// TIA Portal V17 program export: 0 tag tables, 0 data types, 1 data blocks, 1 code blocks (in call order from the OBs), 0 instance data blocks

DATA_BLOCK "流水灯定时器"   // DB1
{ S7_Optimized_Access := 'FALSE' }
   VAR
      黄灯计时 : TON_TIME;
      蓝灯计时 : TON_TIME;
      紫灯计时 : TON_TIME;
      红灯亮计时 : TON_TIME;
      红灯灭计时 : TON_TIME;
   END_VAR
BEGIN
END_DATA_BLOCK

ORGANIZATION_BLOCK "Main"   // OB1, LAD, ProgramCycle
TITLE = 作业6：黄蓝紫流水灯与红灯1Hz闪烁
{ S7_Optimized_Access := 'TRUE' }
// 作业6：黄蓝紫流水灯与红灯1Hz闪烁
// stored: SetENOAutomatically false
   VAR_INPUT
      Initial_Call : Bool;   // Initial call of this OB
      Remanence : Bool;   // =True, if remanent data are available
   END_VAR
BEGIN

REGION Network 1: 启停自锁（停止优先）
   // 按开启动，松开后自锁；关为1时立即停止。开关同时按下，停止优先。
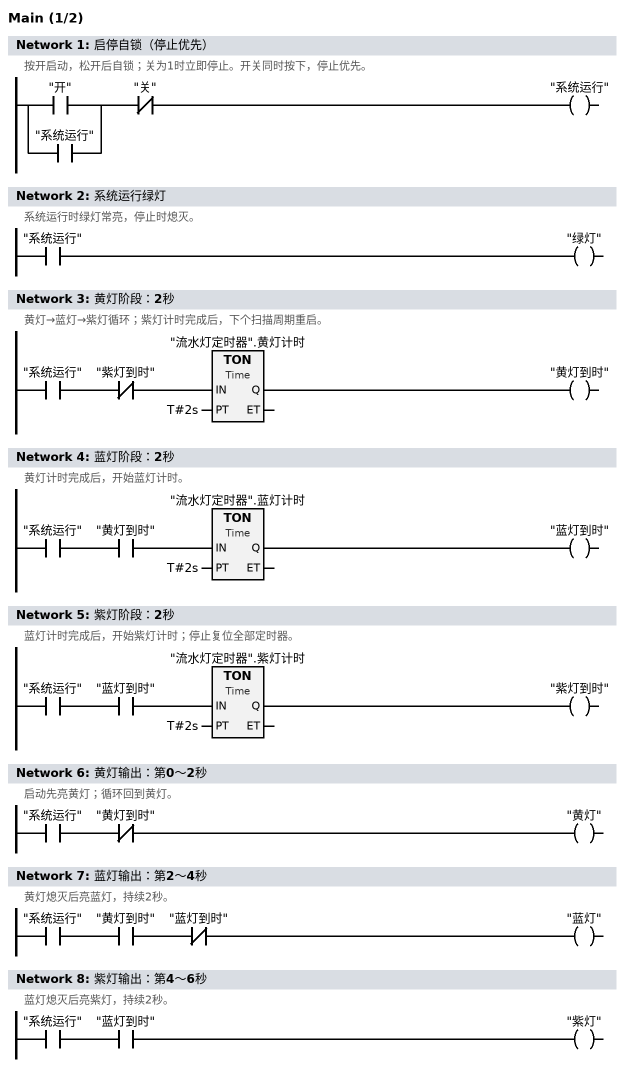
   RUNG wire#powerrail
      Contact( "开" )
      wire#w1
      I_Contact( "关" )
      Coil( "系统运行" )
   END_RUNG
   RUNG wire#powerrail
      Contact( "系统运行" )
   END_RUNG wire#w1
   // the same network as SCL:
   "系统运行" := ("开" OR "系统运行") AND NOT "关";
END_REGION

REGION Network 2: 系统运行绿灯
   // 系统运行时绿灯常亮，停止时熄灭。
   RUNG wire#powerrail
      Contact( "系统运行" )
      Coil( "绿灯" )
   END_RUNG
   // the same network as SCL:
   "绿灯" := "系统运行";
END_REGION

REGION Network 3: 黄灯阶段：2秒
   // 黄灯→蓝灯→紫灯循环；紫灯计时完成后，下个扫描周期重启。
   RUNG wire#powerrail
      Contact( "系统运行" )
      I_Contact( "紫灯到时" )
      { S7_Templates := "time_type := Time" } "流水灯定时器".黄灯计时.TON(pt := T#2s, et =>)
      Coil( "黄灯到时" )
   END_RUNG
   // the same network as SCL:
   "流水灯定时器".黄灯计时.TON(IN := "系统运行" AND NOT "紫灯到时", PT := T#2s);
   "黄灯到时" := "流水灯定时器".黄灯计时.Q;
END_REGION

REGION Network 4: 蓝灯阶段：2秒
   // 黄灯计时完成后，开始蓝灯计时。
   RUNG wire#powerrail
      Contact( "系统运行" )
      Contact( "黄灯到时" )
      { S7_Templates := "time_type := Time" } "流水灯定时器".蓝灯计时.TON(pt := T#2s, et =>)
      Coil( "蓝灯到时" )
   END_RUNG
   // the same network as SCL:
   "流水灯定时器".蓝灯计时.TON(IN := "系统运行" AND "黄灯到时", PT := T#2s);
   "蓝灯到时" := "流水灯定时器".蓝灯计时.Q;
END_REGION

REGION Network 5: 紫灯阶段：2秒
   // 蓝灯计时完成后，开始紫灯计时；停止复位全部定时器。
   RUNG wire#powerrail
      Contact( "系统运行" )
      Contact( "蓝灯到时" )
      { S7_Templates := "time_type := Time" } "流水灯定时器".紫灯计时.TON(pt := T#2s, et =>)
      Coil( "紫灯到时" )
   END_RUNG
   // the same network as SCL:
   "流水灯定时器".紫灯计时.TON(IN := "系统运行" AND "蓝灯到时", PT := T#2s);
   "紫灯到时" := "流水灯定时器".紫灯计时.Q;
END_REGION

REGION Network 6: 黄灯输出：第0～2秒
   // 启动先亮黄灯；循环回到黄灯。
   RUNG wire#powerrail
      Contact( "系统运行" )
      I_Contact( "黄灯到时" )
      Coil( "黄灯" )
   END_RUNG
   // the same network as SCL:
   "黄灯" := "系统运行" AND NOT "黄灯到时";
END_REGION

REGION Network 7: 蓝灯输出：第2～4秒
   // 黄灯熄灭后亮蓝灯，持续2秒。
   RUNG wire#powerrail
      Contact( "系统运行" )
      Contact( "黄灯到时" )
      I_Contact( "蓝灯到时" )
      Coil( "蓝灯" )
   END_RUNG
   // the same network as SCL:
   "蓝灯" := "系统运行" AND "黄灯到时" AND NOT "蓝灯到时";
END_REGION

REGION Network 8: 紫灯输出：第4～6秒
   // 蓝灯熄灭后亮紫灯，持续2秒。
   RUNG wire#powerrail
      Contact( "系统运行" )
      Contact( "蓝灯到时" )
      Coil( "紫灯" )
   END_RUNG
   // the same network as SCL:
   "紫灯" := "系统运行" AND "蓝灯到时";
END_REGION

REGION Network 9: 红灯亮：0.5秒
   // 红灯闪烁周期1秒，亮0.5秒、灭0.5秒。
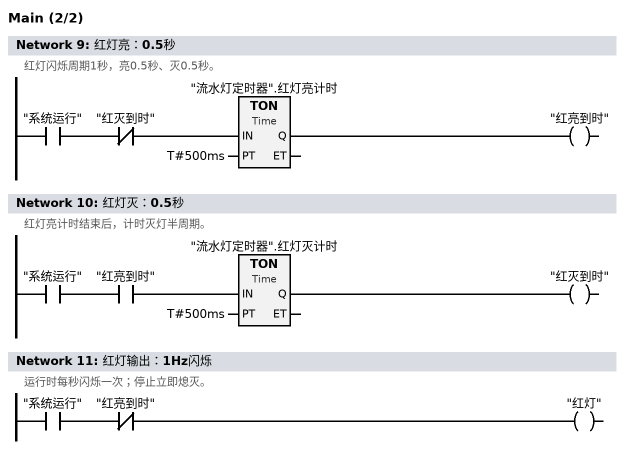
   RUNG wire#powerrail
      Contact( "系统运行" )
      I_Contact( "红灭到时" )
      { S7_Templates := "time_type := Time" } "流水灯定时器".红灯亮计时.TON(pt := T#500ms, et =>)
      Coil( "红亮到时" )
   END_RUNG
   // the same network as SCL:
   "流水灯定时器".红灯亮计时.TON(IN := "系统运行" AND NOT "红灭到时", PT := T#500ms);
   "红亮到时" := "流水灯定时器".红灯亮计时.Q;
END_REGION

REGION Network 10: 红灯灭：0.5秒
   // 红灯亮计时结束后，计时灭灯半周期。
   RUNG wire#powerrail
      Contact( "系统运行" )
      Contact( "红亮到时" )
      { S7_Templates := "time_type := Time" } "流水灯定时器".红灯灭计时.TON(pt := T#500ms, et =>)
      Coil( "红灭到时" )
   END_RUNG
   // the same network as SCL:
   "流水灯定时器".红灯灭计时.TON(IN := "系统运行" AND "红亮到时", PT := T#500ms);
   "红灭到时" := "流水灯定时器".红灯灭计时.Q;
END_REGION

REGION Network 11: 红灯输出：1Hz闪烁
   // 运行时每秒闪烁一次；停止立即熄灭。
   RUNG wire#powerrail
      Contact( "系统运行" )
      I_Contact( "红亮到时" )
      Coil( "红灯" )
   END_RUNG
   // the same network as SCL:
   "红灯" := "系统运行" AND NOT "红亮到时";
END_REGION
END_ORGANIZATION_BLOCK
